// TIA Portal V20 export
DATA_BLOCK "DB_prikazy_tiskarna"   // DB4
{ S7_Optimized_Access := 'TRUE' }
// stored: MemoryReserve 0
   VAR
      task : Array[0..6, 0..255] of Byte;
      DATA : Array[0..255] of Byte;
      ADRESACE_POLE : Int := 1;
      hodnota_pamet : Int := 1;
      cislo_zpravy : Int := 2;   // zpráva má pevný formát mění se pouze číslo které je odesíláno jako string před převedením do stringu je rozseknuto na byte a kopírováno jako jednotlyvý znak
      DATA_RECIVR : Array[0..255] of Byte;
      byte_1 : Byte := 16#30;
      byte_2 : Byte := 16#32;
      text_pole_1 : String[30];   // pole jedno - odkud pochází
      text_pole_2 : String[10];   // pole dvě - datum spotřeby požadovaný formát xx.xx.xxxx
   END_VAR
BEGIN
   task[0,0] := 16#00;   // get_status
   task[0,1..4] := 16#00;
   task[0,5] := 16#06;
   task[0,6] := 16#01;
   task[0,7] := 16#64;
   task[0,8] := 16#00;
   task[0,9] := 16#02;
   task[0,10] := 16#01;
   task[0,11] := 16#45;
   // task[0,255] : get_status
   task[1,0] := 16#00;   // START_TISKU
   task[1,1] := 16#00;   // START_TISKU
   task[1,2] := 16#00;   // START_TISKU
   task[1,3] := 16#00;   // START_TISKU
   task[1,4] := 16#00;   // START_TISKU
   task[1,5] := 16#0D;   // START_TISKU
   task[1,6] := 16#01;   // START_TISKU
   task[1,7] := 16#64;   // START_TISKU
   task[1,8] := 16#00;   // START_TISKU
   task[1,9] := 16#09;   // START_TISKU
   task[1,10] := 16#01;   // START_TISKU
   task[1,11] := 16#20;   // START_TISKU
   task[1,12] := 16#02;   // START_TISKU
   task[1,13] := 16#13;   // START_TISKU
   task[1,14] := 16#00;   // START_TISKU
   task[1,15] := 16#00;   // START_TISKU
   task[1,16] := 16#00;   // START_TISKU
   task[1,17] := 16#00;   // START_TISKU
   task[1,18] := 16#00;   // START_TISKU
   // task[1,255] : START_TISKU
   task[2,0] := 16#00;   // STOP_TISKU
   task[2,1] := 16#00;   // STOP_TISKU
   task[2,2] := 16#00;   // STOP_TISKU
   task[2,3] := 16#00;   // STOP_TISKU
   task[2,4] := 16#00;   // STOP_TISKU
   task[2,5] := 16#0D;   // STOP_TISKU
   task[2,6] := 16#01;   // STOP_TISKU
   task[2,7] := 16#64;   // STOP_TISKU
   task[2,8] := 16#00;   // STOP_TISKU
   task[2,9] := 16#09;   // STOP_TISKU
   task[2,10] := 16#01;   // STOP_TISKU
   task[2,11] := 16#20;   // STOP_TISKU
   task[2,12] := 16#02;   // STOP_TISKU
   task[2,13] := 16#13;   // STOP_TISKU
   task[2,14] := 16#00;   // STOP_TISKU
   task[2,15] := 16#00;   // STOP_TISKU
   task[2,16] := 16#00;   // STOP_TISKU
   task[2,17] := 16#00;   // STOP_TISKU
   task[2,18] := 16#01;   // STOP_TISKU
   // task[2,19] : STOP_TISKU
   // task[2,20] : STOP_TISKU
   // task[2,21] : STOP_TISKU
   task[3,0] := 16#00;
   task[3,1] := 16#00;   // VÝBĚR ZPRÁVY
   task[3,2] := 16#00;   // VÝBĚR ZPRÁVY
   task[3,3] := 16#00;   // VÝBĚR ZPRÁVY
   task[3,4] := 16#00;
   task[3,5] := 16#1A;
   task[3,6] := 16#01;
   task[3,7] := 16#64;
   task[3,8] := 16#00;
   task[3,9] := 16#16;
   task[3,10] := 16#01;
   task[3,11] := 16#20;
   task[3,12] := 16#02;
   task[3,13] := 16#4C;
   task[3,14..18] := 16#00;
   task[3,19] := 16#0C;
   task[3,20] := 16#4D;
   task[3,21] := 16#53;
   task[3,22] := 16#47;
   task[3,23..25] := 16#30;
   task[3,28] := 16#2E;
   task[3,29] := 16#78;
   task[3,30] := 16#6D;
   task[3,31] := 16#6C;
   task[4,0] := 16#00;   // VYPLNĚNÍ DAT MAX 30 ZNAKŮ DO JEDNOHO POLE AKTUÁLNĚ
   task[4,1] := 16#00;   // VYPLNĚNÍ DAT MAX 30 ZNAKŮ DO JEDNOHO POLE AKTUÁLNĚ
   task[4,2] := 16#00;   // VYPLNĚNÍ DAT MAX 30 ZNAKŮ DO JEDNOHO POLE AKTUÁLNĚ
   task[4,3] := 16#00;   // VYPLNĚNÍ DAT MAX 30 ZNAKŮ DO JEDNOHO POLE AKTUÁLNĚ
   task[4,4] := 16#00;   // VYPLNĚNÍ DAT MAX 30 ZNAKŮ DO JEDNOHO POLE AKTUÁLNĚ
   task[4,5] := 16#3C;   // VYPLNĚNÍ DAT MAX 30 ZNAKŮ DO JEDNOHO POLE AKTUÁLNĚ
   task[4,6] := 16#01;   // VYPLNĚNÍ DAT MAX 30 ZNAKŮ DO JEDNOHO POLE AKTUÁLNĚ
   task[4,7] := 16#64;   // VYPLNĚNÍ DAT MAX 30 ZNAKŮ DO JEDNOHO POLE AKTUÁLNĚ
   task[4,8] := 16#00;   // VYPLNĚNÍ DAT MAX 30 ZNAKŮ DO JEDNOHO POLE AKTUÁLNĚ
   task[4,9] := 16#38;   // VYPLNĚNÍ DAT MAX 30 ZNAKŮ DO JEDNOHO POLE AKTUÁLNĚ
   task[4,10] := 16#01;   // VYPLNĚNÍ DAT MAX 30 ZNAKŮ DO JEDNOHO POLE AKTUÁLNĚ
   task[4,11] := 16#CF;   // VYPLNĚNÍ DAT MAX 30 ZNAKŮ DO JEDNOHO POLE AKTUÁLNĚ
   task[4,12] := 16#00;   // VYPLNĚNÍ DAT MAX 30 ZNAKŮ DO JEDNOHO POLE AKTUÁLNĚ
   task[4,13] := 16#00;   // VYPLNĚNÍ DAT MAX 30 ZNAKŮ DO JEDNOHO POLE AKTUÁLNĚ
   task[4,14] := 16#00;   // VYPLNĚNÍ DAT MAX 30 ZNAKŮ DO JEDNOHO POLE AKTUÁLNĚ
   task[4,15] := 16#00;
   task[4,16] := 16#1E;
   task[4,17] := 16#51;
   task[4,18] := 16#57;
   task[4,19] := 16#45;
   task[4,20] := 16#52;
   task[4,21] := 16#54;
   task[4,22] := 16#5A;
   task[4,23] := 16#55;
   task[4,24] := 16#49;
   task[4,25] := 16#4F;
   task[4,26] := 16#50;
   task[4,27] := 16#41;
   task[4,28] := 16#53;
   task[4,29] := 16#44;
   task[4,30] := 16#46;
   task[4,31] := 16#47;
   task[4,32] := 16#48;
   task[4,33] := 16#4A;
   task[4,34] := 16#4B;
   task[4,35] := 16#4C;
   task[4,36] := 16#59;
   task[4,37] := 16#58;
   task[4,38] := 16#43;
   task[4,39] := 16#56;
   task[4,40] := 16#42;
   task[4,41] := 16#4E;
   task[4,42] := 16#4D;
   task[4,43] := 16#31;
   task[4,44] := 16#32;
   task[4,45] := 16#33;
   task[4,46] := 16#34;
   task[4,47..65] := 16#00;
   task[6,0] := 16#00;   // SMAZANÍ A PŘENASTAVENÍ ABY TISKÁRNA NEBAFROVALA ALE TISKLA ODESLANÁ DATA DO KOLA
   task[6,1] := 16#00;   // SMAZANÍ A PŘENASTAVENÍ ABY TISKÁRNA NEBAFROVALA ALE TISKLA ODESLANÁ DATA DO KOLA
   task[6,2] := 16#00;   // SMAZANÍ A PŘENASTAVENÍ ABY TISKÁRNA NEBAFROVALA ALE TISKLA ODESLANÁ DATA DO KOLA
   task[6,3] := 16#00;   // SMAZANÍ A PŘENASTAVENÍ ABY TISKÁRNA NEBAFROVALA ALE TISKLA ODESLANÁ DATA DO KOLA
   task[6,4] := 16#00;   // SMAZANÍ A PŘENASTAVENÍ ABY TISKÁRNA NEBAFROVALA ALE TISKLA ODESLANÁ DATA DO KOLA
   task[6,5] := 16#0D;   // SMAZANÍ A PŘENASTAVENÍ ABY TISKÁRNA NEBAFROVALA ALE TISKLA ODESLANÁ DATA DO KOLA
   task[6,6] := 16#01;   // SMAZANÍ A PŘENASTAVENÍ ABY TISKÁRNA NEBAFROVALA ALE TISKLA ODESLANÁ DATA DO KOLA
   task[6,7] := 16#64;   // SMAZANÍ A PŘENASTAVENÍ ABY TISKÁRNA NEBAFROVALA ALE TISKLA ODESLANÁ DATA DO KOLA
   task[6,8] := 16#00;
   task[6,9] := 16#09;
   task[6,10] := 16#01;
   task[6,11] := 16#CE;
   task[6,12..17] := 16#00;
   task[6,18] := 16#01;
   // DATA_RECIVR[0] : 16#00
   // DATA_RECIVR[1] : 16#00
   // DATA_RECIVR[2] : 16#00
   // DATA_RECIVR[3] : 16#00
   // DATA_RECIVR[4] : 16#00
   // DATA_RECIVR[5] : 16#06
   // DATA_RECIVR[6] : 16#01
   // DATA_RECIVR[7] : 16#64
   // DATA_RECIVR[8] : 16#00
   // DATA_RECIVR[9] : 16#02
   // DATA_RECIVR[10] : 16#01
   // DATA_RECIVR[11] : 16#4F
   // DATA_RECIVR[12] : 16#00
   // DATA_RECIVR[13] : 16#00
   // DATA_RECIVR[14] : 16#00
   // DATA_RECIVR[15] : 16#00
   // DATA_RECIVR[16] : 16#00
   // DATA_RECIVR[17] : 16#06
   // DATA_RECIVR[18] : 16#01
   // DATA_RECIVR[19] : 16#64
   // DATA_RECIVR[20] : 16#00
   // DATA_RECIVR[21] : 16#02
   // DATA_RECIVR[22] : 16#01
   // DATA_RECIVR[23] : 16#4F
   // DATA_RECIVR[24] : 16#00
   // DATA_RECIVR[25] : 16#00
   // DATA_RECIVR[26] : 16#00
   // DATA_RECIVR[27] : 16#00
   // DATA_RECIVR[28] : 16#00
   // DATA_RECIVR[29] : 16#06
   // DATA_RECIVR[30] : 16#01
   // DATA_RECIVR[31] : 16#64
   // DATA_RECIVR[32] : 16#00
   // DATA_RECIVR[33] : 16#02
   // DATA_RECIVR[34] : 16#01
   // DATA_RECIVR[35] : 16#4F
   // DATA_RECIVR[36] : 16#00
   // DATA_RECIVR[37] : 16#00
   // DATA_RECIVR[38] : 16#00
   // DATA_RECIVR[39] : 16#00
   // DATA_RECIVR[40] : 16#00
   // DATA_RECIVR[41] : 16#06
   // DATA_RECIVR[42] : 16#01
   // DATA_RECIVR[43] : 16#64
   // DATA_RECIVR[44] : 16#00
   // DATA_RECIVR[45] : 16#02
   // DATA_RECIVR[46] : 16#01
   // DATA_RECIVR[47] : 16#4F
   // DATA_RECIVR[48] : 16#00
   // DATA_RECIVR[49] : 16#00
   // DATA_RECIVR[50] : 16#00
   // DATA_RECIVR[51] : 16#00
   // DATA_RECIVR[52] : 16#00
   // DATA_RECIVR[53] : 16#06
   // DATA_RECIVR[54] : 16#01
   // DATA_RECIVR[55] : 16#64
   // DATA_RECIVR[56] : 16#00
   // DATA_RECIVR[57] : 16#02
   // DATA_RECIVR[58] : 16#01
   // DATA_RECIVR[59] : 16#4F
   // DATA_RECIVR[60] : 16#00
   // DATA_RECIVR[61] : 16#00
   // DATA_RECIVR[62] : 16#00
   // DATA_RECIVR[63] : 16#00
   // DATA_RECIVR[64] : 16#00
   // DATA_RECIVR[65] : 16#06
   // DATA_RECIVR[66] : 16#01
   // DATA_RECIVR[67] : 16#64
   // DATA_RECIVR[68] : 16#00
   // DATA_RECIVR[69] : 16#02
   // DATA_RECIVR[70] : 16#01
   // DATA_RECIVR[71] : 16#4F
   // DATA_RECIVR[72] : 16#00
   // DATA_RECIVR[73] : 16#00
   // DATA_RECIVR[74] : 16#00
   // DATA_RECIVR[75] : 16#00
   // DATA_RECIVR[76] : 16#00
   // DATA_RECIVR[77] : 16#06
   // DATA_RECIVR[78] : 16#01
   // DATA_RECIVR[79] : 16#64
   // DATA_RECIVR[80] : 16#00
   // DATA_RECIVR[81] : 16#02
   // DATA_RECIVR[82] : 16#01
   // DATA_RECIVR[83] : 16#4F
   // DATA_RECIVR[84] : 16#00
   // DATA_RECIVR[85] : 16#00
   // DATA_RECIVR[86] : 16#00
   // DATA_RECIVR[87] : 16#00
   // DATA_RECIVR[88] : 16#00
   // DATA_RECIVR[89] : 16#06
   // DATA_RECIVR[90] : 16#01
   // DATA_RECIVR[91] : 16#64
   // DATA_RECIVR[92] : 16#00
   // DATA_RECIVR[93] : 16#02
   // DATA_RECIVR[94] : 16#01
   // DATA_RECIVR[95] : 16#4F
   // DATA_RECIVR[96] : 16#00
   // DATA_RECIVR[97] : 16#00
   // DATA_RECIVR[98] : 16#00
   // DATA_RECIVR[99] : 16#00
   // DATA_RECIVR[100] : 16#00
   // DATA_RECIVR[101] : 16#06
   // DATA_RECIVR[102] : 16#01
   // DATA_RECIVR[103] : 16#64
   // DATA_RECIVR[104] : 16#00
   // DATA_RECIVR[105] : 16#02
   // DATA_RECIVR[106] : 16#01
   // DATA_RECIVR[107] : 16#4F
   // DATA_RECIVR[108] : 16#00
   // DATA_RECIVR[109] : 16#00
   // DATA_RECIVR[110] : 16#00
   // DATA_RECIVR[111] : 16#00
   // DATA_RECIVR[112] : 16#00
   // DATA_RECIVR[113] : 16#06
   // DATA_RECIVR[114] : 16#01
   // DATA_RECIVR[115] : 16#64
   // DATA_RECIVR[116] : 16#00
   // DATA_RECIVR[117] : 16#02
   // DATA_RECIVR[118] : 16#01
   // DATA_RECIVR[119] : 16#4F
   // DATA_RECIVR[120] : 16#00
   // DATA_RECIVR[121] : 16#00
   // DATA_RECIVR[122] : 16#00
   // DATA_RECIVR[123] : 16#00
   // DATA_RECIVR[124] : 16#00
   // DATA_RECIVR[125] : 16#06
   // DATA_RECIVR[126] : 16#01
   // DATA_RECIVR[127] : 16#64
   // DATA_RECIVR[128] : 16#00
   // DATA_RECIVR[129] : 16#02
   // DATA_RECIVR[130] : 16#01
   // DATA_RECIVR[131] : 16#4F
   // DATA_RECIVR[132] : 16#00
   // DATA_RECIVR[133] : 16#00
   // DATA_RECIVR[134] : 16#00
   // DATA_RECIVR[135] : 16#00
   // DATA_RECIVR[136] : 16#00
   // DATA_RECIVR[137] : 16#06
   // DATA_RECIVR[138] : 16#01
   // DATA_RECIVR[139] : 16#64
   // DATA_RECIVR[140] : 16#00
   // DATA_RECIVR[141] : 16#02
   // DATA_RECIVR[142] : 16#01
   // DATA_RECIVR[143] : 16#4F
   // DATA_RECIVR[144] : 16#00
   // DATA_RECIVR[145] : 16#00
   // DATA_RECIVR[146] : 16#00
   // DATA_RECIVR[147] : 16#00
   // DATA_RECIVR[148] : 16#00
   // DATA_RECIVR[149] : 16#06
   // DATA_RECIVR[150] : 16#01
   // DATA_RECIVR[151] : 16#64
   // DATA_RECIVR[152] : 16#00
   // DATA_RECIVR[153] : 16#02
   // DATA_RECIVR[154] : 16#01
   // DATA_RECIVR[155] : 16#4F
   // DATA_RECIVR[156] : 16#00
   // DATA_RECIVR[157] : 16#00
   // DATA_RECIVR[158] : 16#00
   // DATA_RECIVR[159] : 16#00
   // DATA_RECIVR[160] : 16#00
   // DATA_RECIVR[161] : 16#06
   // DATA_RECIVR[162] : 16#01
   // DATA_RECIVR[163] : 16#64
   // DATA_RECIVR[164] : 16#00
   // DATA_RECIVR[165] : 16#02
   // DATA_RECIVR[166] : 16#01
   // DATA_RECIVR[167] : 16#4F
   // DATA_RECIVR[168] : 16#00
   // DATA_RECIVR[169] : 16#00
   // DATA_RECIVR[170] : 16#00
   // DATA_RECIVR[171] : 16#00
   // DATA_RECIVR[172] : 16#00
   // DATA_RECIVR[173] : 16#06
   // DATA_RECIVR[174] : 16#01
   // DATA_RECIVR[175] : 16#64
   // DATA_RECIVR[176] : 16#00
   // DATA_RECIVR[177] : 16#02
   // DATA_RECIVR[178] : 16#01
   // DATA_RECIVR[179] : 16#4F
   // DATA_RECIVR[180] : 16#00
   // DATA_RECIVR[181] : 16#00
   // DATA_RECIVR[182] : 16#00
   // DATA_RECIVR[183] : 16#00
   // DATA_RECIVR[184] : 16#00
   // DATA_RECIVR[185] : 16#06
   // DATA_RECIVR[186] : 16#01
   // DATA_RECIVR[187] : 16#64
   // DATA_RECIVR[188] : 16#00
   // DATA_RECIVR[189] : 16#02
   // DATA_RECIVR[190] : 16#01
   // DATA_RECIVR[191] : 16#4F
   // DATA_RECIVR[192] : 16#00
   // DATA_RECIVR[193] : 16#00
   // DATA_RECIVR[194] : 16#00
   // DATA_RECIVR[195] : 16#00
   // DATA_RECIVR[196] : 16#00
   // DATA_RECIVR[197] : 16#06
   // DATA_RECIVR[198] : 16#01
   // DATA_RECIVR[199] : 16#64
   // DATA_RECIVR[200] : 16#00
   // DATA_RECIVR[201] : 16#02
   // DATA_RECIVR[202] : 16#01
   // DATA_RECIVR[203] : 16#4F
   // DATA_RECIVR[204] : 16#00
   // DATA_RECIVR[205] : 16#00
   // DATA_RECIVR[206] : 16#00
   // DATA_RECIVR[207] : 16#00
   // DATA_RECIVR[208] : 16#00
   // DATA_RECIVR[209] : 16#06
   // DATA_RECIVR[210] : 16#01
   // DATA_RECIVR[211] : 16#64
   // DATA_RECIVR[212] : 16#00
   // DATA_RECIVR[213] : 16#02
   // DATA_RECIVR[214] : 16#01
   // DATA_RECIVR[215] : 16#4F
   // DATA_RECIVR[216] : 16#00
   // DATA_RECIVR[217] : 16#00
   // DATA_RECIVR[218] : 16#00
   // DATA_RECIVR[219] : 16#00
   // DATA_RECIVR[220] : 16#00
   // DATA_RECIVR[221] : 16#06
   // DATA_RECIVR[222] : 16#01
   // DATA_RECIVR[223] : 16#64
   // DATA_RECIVR[224] : 16#00
   // DATA_RECIVR[225] : 16#02
   // DATA_RECIVR[226] : 16#01
   // DATA_RECIVR[227] : 16#4F
   // DATA_RECIVR[228] : 16#00
   // DATA_RECIVR[229] : 16#00
   // DATA_RECIVR[230] : 16#00
   // DATA_RECIVR[231] : 16#00
   // DATA_RECIVR[232] : 16#00
   // DATA_RECIVR[233] : 16#07
   // DATA_RECIVR[234] : 16#01
   // DATA_RECIVR[235] : 16#64
   // DATA_RECIVR[236] : 16#00
   // DATA_RECIVR[237] : 16#03
   // DATA_RECIVR[238] : 16#01
   // DATA_RECIVR[239] : 16#31
   // DATA_RECIVR[240] : 16#04
   // DATA_RECIVR[241] : 16#00
   // DATA_RECIVR[242] : 16#00
   // DATA_RECIVR[243] : 16#00
   // DATA_RECIVR[244] : 16#00
   // DATA_RECIVR[245] : 16#00
   // DATA_RECIVR[246] : 16#07
   // DATA_RECIVR[247] : 16#01
   // DATA_RECIVR[248] : 16#64
   // DATA_RECIVR[249] : 16#00
   // DATA_RECIVR[250] : 16#03
   // DATA_RECIVR[251] : 16#01
   // DATA_RECIVR[252] : 16#45
   // DATA_RECIVR[253] : 16#00
   // DATA_RECIVR[254] : 16#00
   // DATA_RECIVR[255] : 16#00
END_DATA_BLOCK
